FUNCTION_BLOCK DEMUX_2 (* Basic Function Block Type *)
  (* Standard: 61499-2 *)
  (* Version 0.0, 10/19/2026, macie, Schneider Electric, Template *)
  PACKAGE Main;
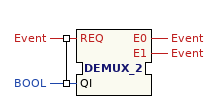
  EVENT_INPUT
    REQ WITH QI; (* Normal Execution Request *)
  END_EVENT
  EVENT_OUTPUT
    E0; (* Execution Confirmation *)
    E1;
  END_EVENT
  VAR_INPUT
    QI : BOOL; (* Input event qualifier *)
  END_VAR
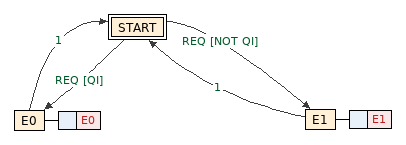
  EC_STATES
    START; (* Initial State *)
    E0 : -> E0; (* Normal execution *)
    E1 : -> E1;
  END_STATES
  EC_TRANSITIONS
    START TO E0 := REQ [QI];
    E0 TO START := 1;
    START TO E1 := REQ [NOT QI];
    E1 TO START := 1;
  END_TRANSITIONS
  ALGORITHM INIT IN ST: (* Initialization algorithm *)
;
  END_ALGORITHM
  ALGORITHM REQ IN ST: (* Normally executed algorithm *)
;
  END_ALGORITHM
END_FUNCTION_BLOCK
